Staubli VAL3: setSpeed.pgx

program setSpeed()
  local bool l_bErr
  local num l_nResult
  local num l_nSpeed
begin
  //设置机器人速度
  if getProfile()=="customer"
    call io:getAnaIO(io:aInput[1],l_nSpeed,l_bErr)
    if l_bErr==false
      l_nSpeed=round(l_nSpeed)
      if l_nSpeed>0 and l_nSpeed<=100 and getMonitorSpeed()!=l_nSpeed
        setMonitorSpeed(l_nSpeed)
      endIf
    endIf
  endIf
  //手动设回default权限
  if workingMode()==4 and getProfile()!="customer"
    l_nResult=setProfile("customer","")
  endIf
  if workingMode()==1 and getProfile()=="customer"
    l_nResult=setProfile("default","")
  endIf
end
